(* IEC 61131-3 sources: codesys-to-s7/tests/corpus/C2S7-POU-INIT/neg, 1 file *)

(* ---- input.st ---- *)
FUNCTION F_Case : INT
VAR_INPUT
    x : BOOL;
END_VAR
VAR_OUTPUT
    o : INT;
END_VAR
o := 1; F_Case := 1;
END_FUNCTION
